{attribute 'qualified_only'}
VAR_GLOBAL
    // Results of the FEM 9.851 double-cycle test, for the performance protocol.
    lrDoubleCycleCalc     : LREAL;   // calculated [s]
    lrDoubleCycleMeasured : LREAL;   // measured in the simulation [s]
    lrDoubleCyclesPerHour : LREAL;   // 3600 / measured
END_VAR

(* stored: Version 1.1.0.1
   GVL GVL_Test: Id {5af14218-5507-4eeb-b5e5-176a038ccb51} *)
